(* PLC project PR_StackUltraWeldSeq_Soft2_PLC, SiemensToBackhoff Siemens TIA Portal → Beckhoff TwinCAT PLCopen Converter 2.2 *)
(* stored: creationDateTime 2026-10-12T09:25:18.517675, modificationDateTime 2026-10-12T09:25:18.517675 *)

FUNCTION_BLOCK PR_StackUltraWeldSeq_Soft2
VAR_INPUT
	iAbort : BOOL;
	iAutoRunning : BOOL;
	iFaultReset : BOOL;
	iPartClampClose : BOOL;
	iPartClampOpen : BOOL;
	iPartNotWorkable : BOOL;
	iPartWorkable : BOOL;
	iRFReadDone : BOOL;
	iRFReadError : BOOL;
	iRFWriteDone : BOOL;
	iRFWriteError : BOOL;
	iReject : BOOL;
	iReset_fault : BOOL;
	iRetry : BOOL;
	iRetryCount : INT;
	iSstMode : BOOL;
	iSstPB : BOOL;
	iStartFrmFibroseq : BOOL;
	iWeldComplete : BOOL;
	iWeldTabDown : BOOL;
	iWeldTabUp : BOOL;
	iStartFrmFibroSeq_1 : BOOL;
	iAutorunning_1 : BOOL;
END_VAR
VAR_OUTPUT
	qError : ARRAY[0..3] OF BOOL;
	qFumeExtractorON : BOOL;
	qMessage : ARRAY[0..2] OF BOOL;
	qPartClampClose : BOOL;
	qPartClampOpen : BOOL;
	qStackUltraWeldOver : BOOL;
	qWeldTabDown : BOOL;
	qWeldTabUp : BOOL;
END_VAR
VAR
	c20_ChkRecovery_T1 : BOOL;
	c20_ChkRecovery_T2 : BOOL;
	c20_ChkRecovery_T3 : BOOL;
	c21_WtRFIDReadOver_T1 : BOOL;
	c21_WtRFIDReadOver_T2 : BOOL;
	c22_ChkReadRetryCnt_T1 : BOOL;
	c22_ChkReadRetryCnt_T2 : BOOL;
	c23_ChkPartWrkSts_T1 : BOOL;
	c23_ChkPartWrkSts_T2 : BOOL;
	c24_WtOpDecision_T1 : BOOL;
	c24_WtOpDecision_T2 : BOOL;
	c81_WtRFIDWriteOver_T1 : BOOL;
	c81_WtRFIDWriteOver_T2 : BOOL;
	c82_ChkWriteRetryCnt_T1 : BOOL;
	c82_ChkWriteRetryCnt_T2 : BOOL;
	c83_WtOpDecisionWrite_T1 : BOOL;
	c83_WtOpDecisionWrite_T2 : BOOL;
	StateNo : INT;
	s10_WtStartFrmFibro : BOOL;
	s10_WtStartFrmFibro_T1 : BOOL;
	s1_WtResetRel : BOOL;
	s1_WtResetRel_T1 : BOOL;
	s20_ChkRecovery : BOOL;
	s20_ChkRecovery_T1 : BOOL;
	s20_ChkRecovery_T2 : BOOL;
	s20_ChkRecovery_T3 : BOOL;
	s21_WtRFIDReadOver : BOOL;
	s21_WtRFIDReadOver_T1 : BOOL;
	s21_WtRFIDReadOver_T2 : BOOL;
	s22_ChkReadRetryCnt : BOOL;
	s22_ChkReadRetryCnt_T1 : BOOL;
	s22_ChkReadRetryCnt_T2 : BOOL;
	s23_ChkPartWrkSts : BOOL;
	s23_ChkPartWrkSts_T1 : BOOL;
	s23_ChkPartWrkSts_T2 : BOOL;
	s24_WtOpDecision : BOOL;
	s24_WtOpDecision_T1 : BOOL;
	s24_WtOpDecision_T2 : BOOL;
	s30_WtOpAck : BOOL;
	s30_WtOpAck_T1 : BOOL;
	s40_WtPartClamp : BOOL;
	s40_WtPartClamp_T1 : BOOL;
	s50_WtWeldTabDown : BOOL;
	s50_WtWeldTabDown_T1 : BOOL;
	s60_WtWeldComplete : BOOL;
	s60_WtWeldComplete_T1 : BOOL;
	s70_WtWeldTabUp : BOOL;
	s70_WtWeldTabUp_T1 : BOOL;
	s80_WtPartClampOpen : BOOL;
	s80_WtPartClampOpen_T1 : BOOL;
	s81_WtRFIDWriteOver : BOOL;
	s81_WtRFIDWriteOver_T1 : BOOL;
	s81_WtRFIDWriteOver_T2 : BOOL;
	s82_ChkWriteRetryCnt : BOOL;
	s82_ChkWriteRetryCnt_T1 : BOOL;
	s82_ChkWriteRetryCnt_T2 : BOOL;
	s83_WtOpDecisionWrite : BOOL;
	s83_WtOpDecisionWrite_T1 : BOOL;
	s83_WtOpDecisionWrite_T2 : BOOL;
	s90_WtStartLow : BOOL;
	s90_WtStartLow_T1 : BOOL;
	sRFReadRetryCount : INT;
	sRFWriteRetryCount : INT;
	sSst : BOOL;
	sSstPulse : BOOL;
	sSstRise : R_TRIG;
	sStWtResetRel : BOOL;
	sStWtResetRel_T1 : BOOL;
	sWeldDlyOver : BOOL;
	sweldingInProgress : INT;
	SET : BOOL;
	c20_ChkRecovery_clamp : BOOL;
END_VAR
VAR_TEMP
	tOne : BOOL;
	tRFReadRetryCountInc : INT;
	tRFWriteRetryCountInc : INT;
END_VAR
  VAR  (* added by the conversion: wires and edge detectors of the diagram *)
    _w24 : BOOL;
    _w26 : BOOL;
    _w39 : BOOL;
    _w41 : BOOL;
    _w42 : BOOL;
    _w59 : BOOL;
    _w62 : BOOL;
    _w63 : BOOL;
    _w109 : BOOL;
    _w112 : BOOL;
    _w113 : BOOL;
    _w114 : BOOL;
    _w115 : BOOL;
    _w128 : BOOL;
    _w130 : BOOL;
    _w131 : BOOL;
    _w162 : BOOL;
    _w165 : BOOL;
    _w166 : BOOL;
    _w167 : BOOL;
    _w195 : BOOL;
    _w197 : BOOL;
    _w198 : BOOL;
    _w199 : BOOL;
    _w223 : BOOL;
    _w226 : BOOL;
    _w227 : BOOL;
    _w228 : BOOL;
    _w249 : BOOL;
    _w251 : BOOL;
    _w252 : BOOL;
    _w253 : BOOL;
    _w266 : BOOL;
    _w268 : BOOL;
    _w269 : BOOL;
    _w290 : BOOL;
    _w292 : BOOL;
    _w293 : BOOL;
    _w310 : BOOL;
    _w313 : BOOL;
    _w314 : BOOL;
    _w333 : BOOL;
    _w337 : BOOL;
    _w338 : BOOL;
    _w355 : BOOL;
    _w357 : BOOL;
    _w358 : BOOL;
    _w386 : BOOL;
    _w390 : BOOL;
    _w391 : BOOL;
    _w392 : BOOL;
    _w424 : BOOL;
    _w426 : BOOL;
    _w427 : BOOL;
    _w428 : BOOL;
    _w457 : BOOL;
    _w459 : BOOL;
    _w460 : BOOL;
    _w461 : BOOL;
    _w474 : BOOL;
    _w477 : BOOL;
    _w478 : BOOL;
  END_VAR

(* LD diagram, written out as Structured Text *)
(* Network 1 *)
(* Create Single Step Pulse bit *)
(* Create Single Step bit *)
(* Transition for STATE Num:0 Reset Released *)
(* STATE Num:0 Reset Released *)
(* Transition for STATE Num:1 Wait for Rest Release *)
(* STATE Num:1 Wait for Rest Release *)
(* Transition for STATE Num:10 Wait for Start From Fibro Main seq *)
(* STATE Num:10 Wait for Start From Fibro Main seq *)
(* Condition1 for STATE Num:20 Check Recovery //Human in Loop required *)
(* Condition for STATE Num:20 Check Recovery clamp branch *)
(* Condition2 for STATE Num:20 Check Recovery *)
(* Condition3 for STATE Num:20 Check Recovery *)
(* Transition for STATE Num:20 Check Recovery *)
(* STATE Num:20 Check Recovery *)
(* Transition for STATE Num:30 Wait for Operator Ack *)
(* STATE Num:30 Wait for Operator Ack *)
(* Actions for STATE Num:30 Wait for Operator Ack - qError[0] := 1 *)
(* Condition1 for STATE Num:21 Wait For RFID Read Over *)
(* Condition2 for STATE Num:21 Wait For RFID Read Over *)
(* Transition for STATE Num:21 Wait For RFID Read Over *)
(* STATE Num:21 Wait For RFID Read Over *)
(* Condition1 for STATE Num:22 Check Read Retry Count Over *)
(* Condition2 for STATE Num:22 Check Read Retry Count Over *)
(* Transition for STATE Num:22 Check Read Retry Count Over *)
(* STATE Num:22 Check Read Retry Count Over *)
(* Condition1 for STATE Num:23 Check Part Workable Status *)
(* Condition2 for STATE Num:23 Check Part Workable Status *)
(* Transition for STATE Num:23 Check Part Workable Status *)
(* STATE Num:23 Check Part Workable Status *)
(* Actions for STATE Num:23 T1 - qMessage[2] := 1 *)
(* Transition for STATE Num:24 Wait For Operator Decision_Read *)
(* STATE Num:24 Wait For Operator Decision_Read *)
(* Transition for STATE Num:40 Wait for Part Clamp *)
(* STATE Num:40 Wait for Part Clamp *)
(* Actions for STATE Num:40 Wait for Part Clamp - qPartClampClose := 1 *)
(* Actions for STATE Num:40 Wait for Part Clamp - qFumeExtractorON := 1 *)
(* Transition for STATE Num:50 Wait for Weld Tab Down *)
(* STATE Num:50 Wait for Weld Tab Down *)
(* Actions for STATE Num:50 Wait for Weld Tab Down - qWeldTabDown := 1 *)
(* Transition for STATE Num:60 Wait for Weld Complete *)
(* STATE Num:60 Wait for Weld Complete *)
(* Actions for STATE Num:60 Wait for Weld Complete - if !iWeldComplete & sWeldDlyOver Then qError[1]:=1 *)
(* Transition for STATE Num:70 Wait for Weld Tab Up *)
(* STATE Num:70 Wait for Weld Tab Up *)
(* Actions for STATE Num:70 Wait for Weld Tab Up - qWeldTabUp := 1 *)
(* Transition for STATE Num:80 Wait for Part Clamp Open *)
(* STATE Num:80 Wait for Part Clamp Open *)
(* Actions for STATE Num:80 Wait for Part Clamp Open - qPartClampOpen := 1 *)
(* Condition1 for STATE Num:81 Wait For RFID write Over *)
(* Condition2 for STATE Num:81 Wait For RFID write Over *)
(* Transition for STATE Num:81 Wait For RFID write Over *)
(* STATE Num:81 Wait For RFID write Over *)
(* Actions for STATE Num:81 Wait For RFID write Over - qMessage[1] := 1 *)
(* Condition1 for STATE Num:82 Check RFID Write Retry Count Over *)
(* Condition2 for STATE Num:82 Check RFID Write Retry Count Over *)
(* Transition for STATE Num:82 Check RFID Write Retry Count Over *)
(* STATE Num:82 Check RFID Write Retry Count Over *)
(* Actions for STATE Num:82 T1 - qError[3] := 1 *)
(* Condition1 for STATE Num:83 Wait For Operator Decision_Write *)
(* Condition2 for STATE Num:83 Wait For Operator Decision_Write *)
(* Transition for STATE Num:83 Wait For Operator Decision_Write *)
(* STATE Num:83 Wait For Operator Decision_Write *)
(* Transition for STATE Num:90 Wait For Start Low *)
(* STATE Num:90 Wait For Start Low *)
(* Actions for STATE Num:90 Wait For Start Low - qStackUltraWeldOver := 1 *)
(* Actions for STATE Num:60 Wait for Weld Complete - sweldingInProgress := 1 *)
(* Actions for STATE Num:80 Wait for Part Clamp Open - qFumeExtractorON := 0 *)
(* Actions for STATE Num:81 Wait For RFID write Over - sRFWriteRetryCount increment *)
(* Actions for STATE Num:21 T1/T2 - qMessage[0] := 1 and sRFReadRetryCount increment *)
(* Actions for STATE Num:22 T1 - qError[2] := 1/Actions for STATE Num:83 Wait For Operator Decision_Write - qError[2] := 1 *)
tOne := tOne OR NOT tOne;
sSstRise(CLK := iSstPB);
sSstPulse := sSstRise.Q;
sSst := iSstMode AND sSstPulse OR NOT iSstMode;
sStWtResetRel_T1 := sStWtResetRel AND iAutoRunning;
_w24 := sStWtResetRel;
_w26 := (_w24 OR NOT iAutoRunning) AND NOT sStWtResetRel_T1;
sStWtResetRel := _w26;
IF _w26 THEN StateNo := 0; END_IF;
s1_WtResetRel_T1 := s1_WtResetRel AND NOT sStWtResetRel AND sSst AND iAutoRunning;
_w39 := s1_WtResetRel;
_w41 := (_w39 OR sStWtResetRel_T1) AND NOT sStWtResetRel;
_w42 := _w41 AND NOT s1_WtResetRel_T1;
s1_WtResetRel := _w42;
IF _w42 THEN StateNo := 1; END_IF;
s10_WtStartFrmFibro_T1 := s10_WtStartFrmFibro AND NOT sStWtResetRel AND sSst AND iStartFrmFibroseq;
IF s10_WtStartFrmFibro AND NOT sStWtResetRel AND sSst AND iStartFrmFibroseq THEN sRFReadRetryCount := 0; END_IF;
IF s10_WtStartFrmFibro AND NOT sStWtResetRel AND sSst AND iStartFrmFibroseq THEN sRFWriteRetryCount := 0; END_IF;
_w59 := s10_WtStartFrmFibro;
_w62 := (_w59 OR s1_WtResetRel_T1 OR s90_WtStartLow_T1) AND NOT sStWtResetRel;
_w63 := _w62 AND NOT s10_WtStartFrmFibro_T1;
s10_WtStartFrmFibro := _w63;
IF _w63 THEN StateNo := 10; END_IF;
c20_ChkRecovery_T1 := sweldingInProgress <> 0 AND c20_ChkRecovery_clamp;
c20_ChkRecovery_clamp := NOT iPartClampClose OR iWeldTabDown;
c20_ChkRecovery_T2 := sweldingInProgress <> 0 AND iPartClampClose AND iWeldTabDown;
c20_ChkRecovery_T3 := sweldingInProgress = 0;
s20_ChkRecovery_T1 := s20_ChkRecovery AND NOT sStWtResetRel AND sSst AND c20_ChkRecovery_T1;
s20_ChkRecovery_T2 := s20_ChkRecovery AND NOT sStWtResetRel AND sSst AND NOT s20_ChkRecovery_T1 AND c20_ChkRecovery_T2;
s20_ChkRecovery_T3 := s20_ChkRecovery AND NOT sStWtResetRel AND sSst AND NOT s20_ChkRecovery_T1 AND NOT s20_ChkRecovery_T1 AND NOT s20_ChkRecovery_T2 AND c20_ChkRecovery_T3;
_w109 := s20_ChkRecovery;
_w112 := (_w109 OR s10_WtStartFrmFibro_T1 OR s30_WtOpAck_T1) AND NOT sStWtResetRel;
_w113 := _w112 AND NOT s20_ChkRecovery_T1;
_w114 := _w113 AND NOT s20_ChkRecovery_T2;
_w115 := _w114 AND NOT s20_ChkRecovery_T3;
s20_ChkRecovery := _w115;
IF _w115 THEN StateNo := 20; END_IF;
s30_WtOpAck_T1 := s30_WtOpAck AND NOT sStWtResetRel AND sSst AND iFaultReset;
_w128 := s30_WtOpAck;
_w130 := (_w128 OR s20_ChkRecovery_T1) AND NOT sStWtResetRel;
_w131 := _w130 AND NOT s30_WtOpAck_T1;
s30_WtOpAck := _w131;
IF _w131 THEN StateNo := 30; END_IF;
qError[0] := s30_WtOpAck;
c21_WtRFIDReadOver_T1 := iRFReadError;
c21_WtRFIDReadOver_T2 := iRFReadDone;
s21_WtRFIDReadOver_T1 := s21_WtRFIDReadOver AND NOT sStWtResetRel AND sSst AND c21_WtRFIDReadOver_T1;
IF s21_WtRFIDReadOver AND NOT sStWtResetRel AND sSst AND c21_WtRFIDReadOver_T1 THEN sRFReadRetryCount := sRFReadRetryCount + 1; END_IF;
s21_WtRFIDReadOver_T2 := s21_WtRFIDReadOver AND NOT sStWtResetRel AND sSst AND NOT s21_WtRFIDReadOver_T1 AND c21_WtRFIDReadOver_T2;
_w162 := s21_WtRFIDReadOver;
_w165 := (_w162 OR s20_ChkRecovery_T3 OR s24_WtOpDecision_T2) AND NOT sStWtResetRel;
_w166 := _w165 AND NOT s21_WtRFIDReadOver_T1;
_w167 := _w166 AND NOT s21_WtRFIDReadOver_T2;
s21_WtRFIDReadOver := _w167;
IF _w167 THEN StateNo := 21; END_IF;
c22_ChkReadRetryCnt_T1 := sRFReadRetryCount > iRetryCount;
c22_ChkReadRetryCnt_T2 := sRFReadRetryCount <= iRetryCount;
s22_ChkReadRetryCnt_T1 := s22_ChkReadRetryCnt AND NOT sStWtResetRel AND sSst AND c22_ChkReadRetryCnt_T1;
s22_ChkReadRetryCnt_T2 := s22_ChkReadRetryCnt AND NOT sStWtResetRel AND sSst AND NOT s22_ChkReadRetryCnt_T1 AND c22_ChkReadRetryCnt_T2;
_w195 := s22_ChkReadRetryCnt;
_w197 := (_w195 OR s21_WtRFIDReadOver_T1) AND NOT sStWtResetRel;
_w198 := _w197 AND NOT s22_ChkReadRetryCnt_T1;
_w199 := _w198 AND NOT s22_ChkReadRetryCnt_T2;
s22_ChkReadRetryCnt := _w199;
IF _w199 THEN StateNo := 22; END_IF;
c23_ChkPartWrkSts_T1 := iPartNotWorkable;
c23_ChkPartWrkSts_T2 := iPartWorkable;
s23_ChkPartWrkSts_T1 := s23_ChkPartWrkSts AND NOT sStWtResetRel AND sSst AND c23_ChkPartWrkSts_T1;
s23_ChkPartWrkSts_T2 := s23_ChkPartWrkSts AND NOT sStWtResetRel AND sSst AND NOT s23_ChkPartWrkSts_T1 AND c23_ChkPartWrkSts_T2;
_w223 := s23_ChkPartWrkSts;
_w226 := (_w223 OR s22_ChkReadRetryCnt_T2 OR s21_WtRFIDReadOver_T2) AND NOT sStWtResetRel;
_w227 := _w226 AND NOT s23_ChkPartWrkSts_T1;
_w228 := _w227 AND NOT s23_ChkPartWrkSts_T2;
s23_ChkPartWrkSts := _w228;
IF _w228 THEN StateNo := 23; END_IF;
qMessage[2] := s23_ChkPartWrkSts_T1;
s24_WtOpDecision_T1 := s24_WtOpDecision AND NOT sStWtResetRel AND sSst AND (iReject OR iAbort);
s24_WtOpDecision_T2 := s24_WtOpDecision AND NOT sStWtResetRel AND sSst AND NOT s24_WtOpDecision_T1 AND iRetry;
_w249 := s24_WtOpDecision;
_w251 := (_w249 OR s22_ChkReadRetryCnt_T1) AND NOT sStWtResetRel;
_w252 := _w251 AND NOT s24_WtOpDecision_T1;
_w253 := _w252 AND NOT s24_WtOpDecision_T2;
s24_WtOpDecision := _w253;
IF _w253 THEN StateNo := 24; END_IF;
s40_WtPartClamp_T1 := s40_WtPartClamp AND NOT sStWtResetRel AND sSst AND iPartClampClose;
_w266 := s40_WtPartClamp;
_w268 := (_w266 OR s23_ChkPartWrkSts_T2) AND NOT sStWtResetRel;
_w269 := _w268 AND NOT s40_WtPartClamp_T1;
s40_WtPartClamp := _w269;
IF _w269 THEN StateNo := 40; END_IF;
qPartClampClose := s40_WtPartClamp;
qFumeExtractorON := s40_WtPartClamp;
s50_WtWeldTabDown_T1 := s50_WtWeldTabDown AND NOT sStWtResetRel AND sSst AND iWeldTabDown;
_w290 := s50_WtWeldTabDown;
_w292 := (_w290 OR s40_WtPartClamp_T1) AND NOT sStWtResetRel;
_w293 := _w292 AND NOT s50_WtWeldTabDown_T1;
s50_WtWeldTabDown := _w293;
IF _w293 THEN StateNo := 50; END_IF;
qWeldTabDown := s50_WtWeldTabDown;
s60_WtWeldComplete_T1 := s60_WtWeldComplete AND NOT sStWtResetRel AND sSst AND iWeldComplete;
_w310 := s60_WtWeldComplete;
_w313 := (_w310 OR s20_ChkRecovery_T2 OR s50_WtWeldTabDown_T1) AND NOT sStWtResetRel;
_w314 := _w313 AND NOT s60_WtWeldComplete_T1;
s60_WtWeldComplete := _w314;
IF _w314 THEN StateNo := 60; END_IF;
qError[1] := s60_WtWeldComplete AND NOT iWeldComplete AND sWeldDlyOver;
s70_WtWeldTabUp_T1 := s70_WtWeldTabUp AND NOT sStWtResetRel AND sSst AND iWeldTabUp;
_w333 := s70_WtWeldTabUp;
_w337 := (_w333 OR s60_WtWeldComplete_T1 OR s24_WtOpDecision_T1 OR s23_ChkPartWrkSts_T1) AND NOT sStWtResetRel;
_w338 := _w337 AND NOT s70_WtWeldTabUp_T1;
s70_WtWeldTabUp := _w338;
IF _w338 THEN StateNo := 70; END_IF;
qWeldTabUp := s70_WtWeldTabUp;
s80_WtPartClampOpen_T1 := s80_WtPartClampOpen AND NOT sStWtResetRel AND sSst AND iPartClampOpen;
_w355 := s80_WtPartClampOpen;
_w357 := (_w355 OR s70_WtWeldTabUp_T1) AND NOT sStWtResetRel;
_w358 := _w357 AND NOT s80_WtPartClampOpen_T1;
s80_WtPartClampOpen := _w358;
IF _w358 THEN StateNo := 80; END_IF;
qPartClampOpen := s80_WtPartClampOpen;
c81_WtRFIDWriteOver_T1 := iRFWriteError;
c81_WtRFIDWriteOver_T2 := iRFWriteDone;
s81_WtRFIDWriteOver_T1 := s81_WtRFIDWriteOver AND NOT sStWtResetRel AND sSst AND c81_WtRFIDWriteOver_T1;
s81_WtRFIDWriteOver_T2 := s81_WtRFIDWriteOver AND NOT sStWtResetRel AND sSst AND NOT s81_WtRFIDWriteOver_T1 AND c81_WtRFIDWriteOver_T2;
_w386 := s81_WtRFIDWriteOver;
_w390 := (_w386 OR s80_WtPartClampOpen_T1 OR s82_ChkWriteRetryCnt_T2 OR s83_WtOpDecisionWrite_T2) AND NOT sStWtResetRel;
_w391 := _w390 AND NOT s81_WtRFIDWriteOver_T1;
_w392 := _w391 AND NOT s81_WtRFIDWriteOver_T2;
s81_WtRFIDWriteOver := _w392;
IF _w392 THEN StateNo := 81; END_IF;
qMessage[1] := s81_WtRFIDWriteOver;
c82_ChkWriteRetryCnt_T1 := sRFWriteRetryCount > iRetryCount;
c82_ChkWriteRetryCnt_T2 := sRFWriteRetryCount <= iRetryCount;
s82_ChkWriteRetryCnt_T1 := s82_ChkWriteRetryCnt AND NOT sStWtResetRel AND sSst AND c82_ChkWriteRetryCnt_T1;
s82_ChkWriteRetryCnt_T2 := s82_ChkWriteRetryCnt AND NOT sStWtResetRel AND sSst AND NOT s82_ChkWriteRetryCnt_T1 AND c82_ChkWriteRetryCnt_T2;
_w424 := s82_ChkWriteRetryCnt;
_w426 := (_w424 OR s81_WtRFIDWriteOver_T1) AND NOT sStWtResetRel;
_w427 := _w426 AND NOT s82_ChkWriteRetryCnt_T1;
_w428 := _w427 AND NOT s82_ChkWriteRetryCnt_T2;
s82_ChkWriteRetryCnt := _w428;
IF _w428 THEN StateNo := 82; END_IF;
qError[3] := s82_ChkWriteRetryCnt_T1;
c83_WtOpDecisionWrite_T1 := iReject OR iAbort;
c83_WtOpDecisionWrite_T2 := iRetry;
s83_WtOpDecisionWrite_T1 := s83_WtOpDecisionWrite AND NOT sStWtResetRel AND sSst AND c83_WtOpDecisionWrite_T1;
s83_WtOpDecisionWrite_T2 := s83_WtOpDecisionWrite AND NOT sStWtResetRel AND sSst AND NOT s83_WtOpDecisionWrite_T1 AND c83_WtOpDecisionWrite_T2;
_w457 := s83_WtOpDecisionWrite;
_w459 := (_w457 OR s82_ChkWriteRetryCnt_T1) AND NOT sStWtResetRel;
_w460 := _w459 AND NOT s83_WtOpDecisionWrite_T1;
_w461 := _w460 AND NOT s83_WtOpDecisionWrite_T2;
s83_WtOpDecisionWrite := _w461;
IF _w461 THEN StateNo := 83; END_IF;
s90_WtStartLow_T1 := s90_WtStartLow AND NOT sStWtResetRel AND sSst AND NOT iStartFrmFibroseq;
_w474 := s90_WtStartLow;
_w477 := (_w474 OR s83_WtOpDecisionWrite_T1 OR s81_WtRFIDWriteOver_T2) AND NOT sStWtResetRel;
_w478 := _w477 AND NOT s90_WtStartLow_T1;
s90_WtStartLow := _w478;
IF _w478 THEN StateNo := 90; END_IF;
qStackUltraWeldOver := s90_WtStartLow;
IF s60_WtWeldComplete AND NOT iWeldComplete AND sWeldDlyOver THEN sweldingInProgress := 1; END_IF;
IF s80_WtPartClampOpen THEN qFumeExtractorON := FALSE; END_IF;
IF s81_WtRFIDWriteOver THEN sRFWriteRetryCount := sRFWriteRetryCount + 1; END_IF;
qMessage[0] := s21_WtRFIDReadOver_T1 OR s21_WtRFIDReadOver_T2;
qError[2] := s22_ChkReadRetryCnt_T1 OR s83_WtOpDecisionWrite;
END_FUNCTION_BLOCK
